{attribute 'qualified_only'}
VAR_GLOBAL
	bEnable : BOOL;
	bInputSignal AT %I* : BOOL;
	nCount : UINT := 2;
	nCycleCount : UDINT;
	fValue : LREAL := 1.5;
	sText : STRING := 'fixture';
	aNames : ARRAY[0..3] OF STRING(20) := ['alpha', 'beta', 'gamma', 'delta'];
END_VAR

(* stored: Version 1.1.0.1
   GVL GVL_Fixture: Id {7a37ae27-a581-4317-a77f-629d6dddcc26} *)
